// CFC twin of T_SafeConnShutdown_Tests: the same tests drawn as CFC diagrams, the way a TwinSAFE project is authored.
    FUNCTION_BLOCK T_SafeConnShutdown_Tests_CFC EXTENDS T_SafeCfcTestSuite
    VAR
    // Test_DeactivateShutsDownConnection
    group_1 : T_SafeGroup;
    conn_1 : T_SafeConnection(group := group_1);
    fb_1 : T_SafeConnShutdown(group := group_1, connection := conn_1);
END_VAR

Test_DeactivateShutsDownConnection();

METHOD PRIVATE Test_DeactivateShutsDownConnection
// note: this text did not pass the execution check against the stored diagram
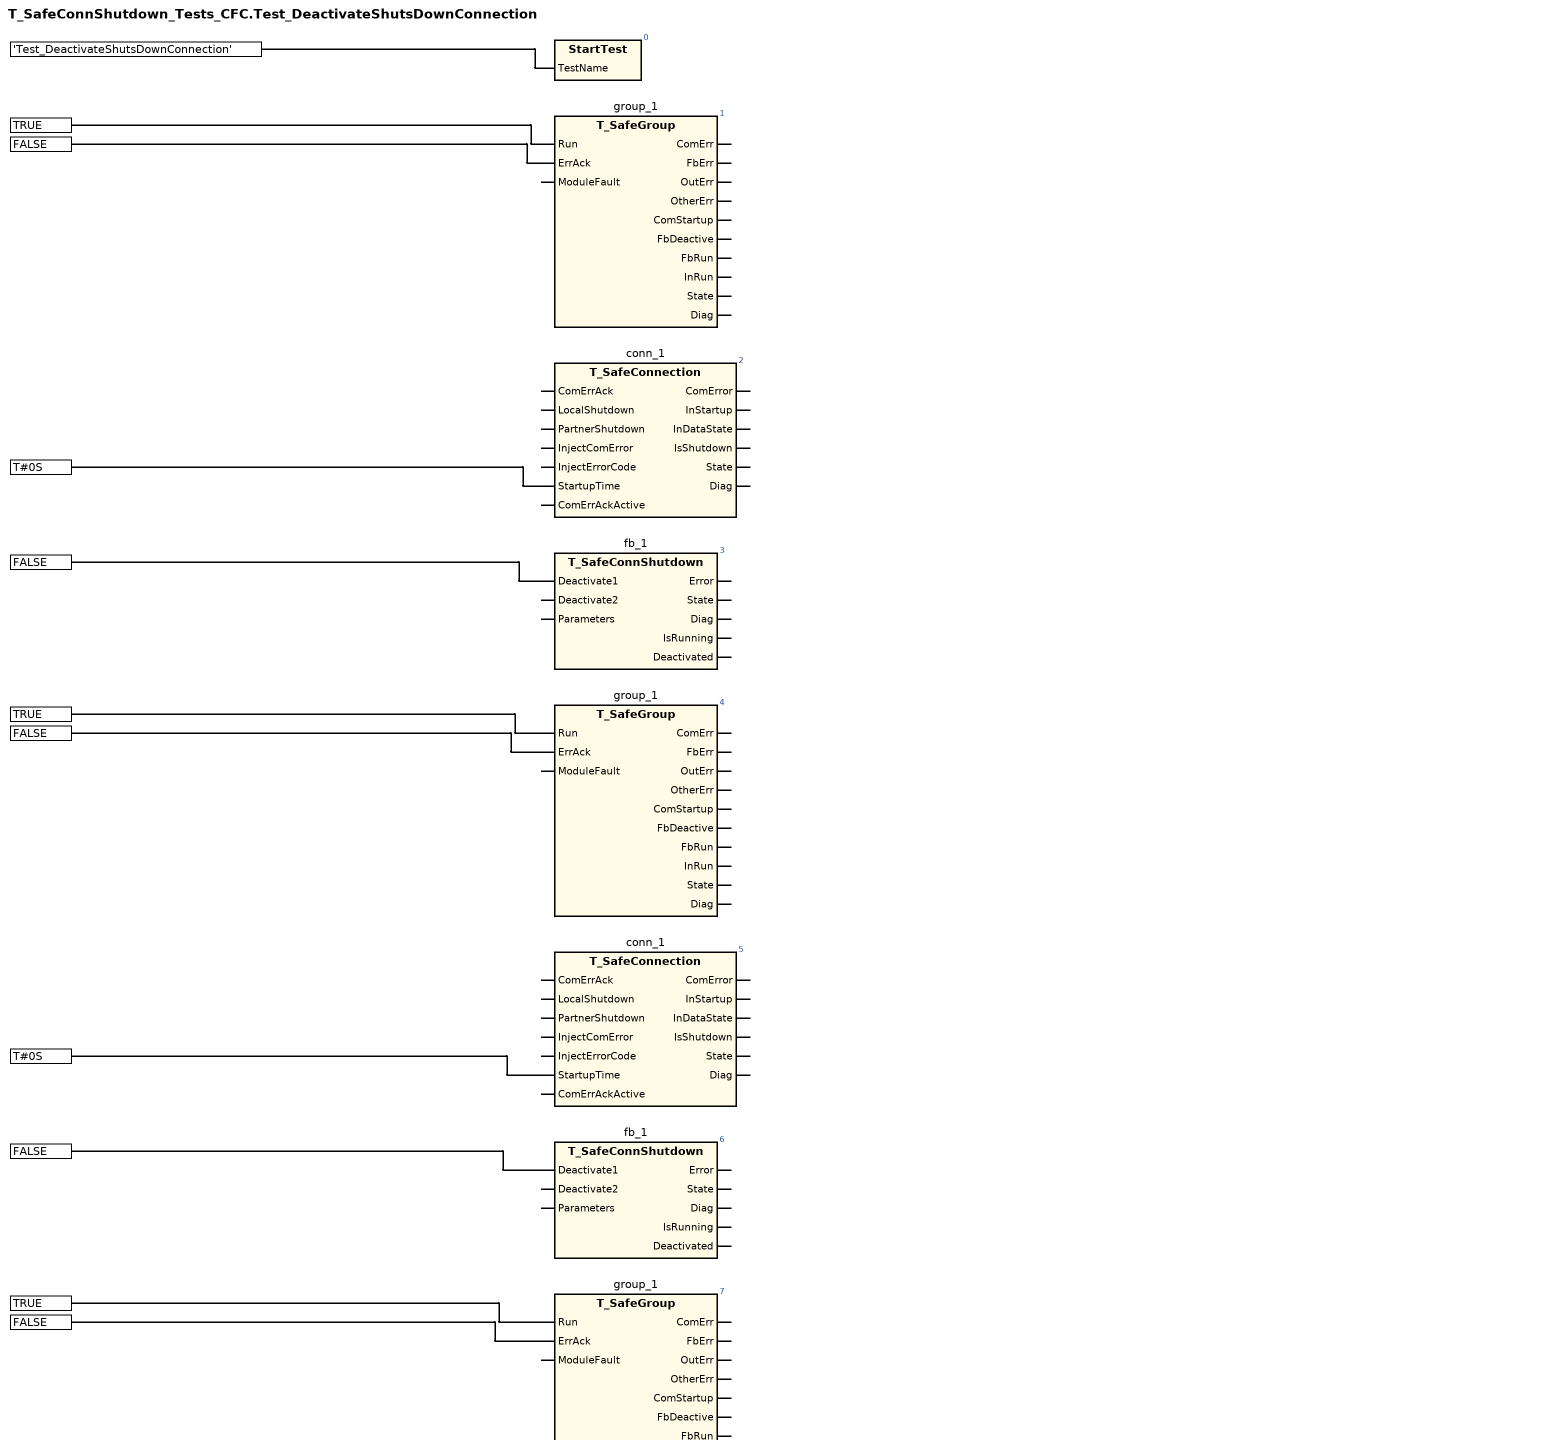
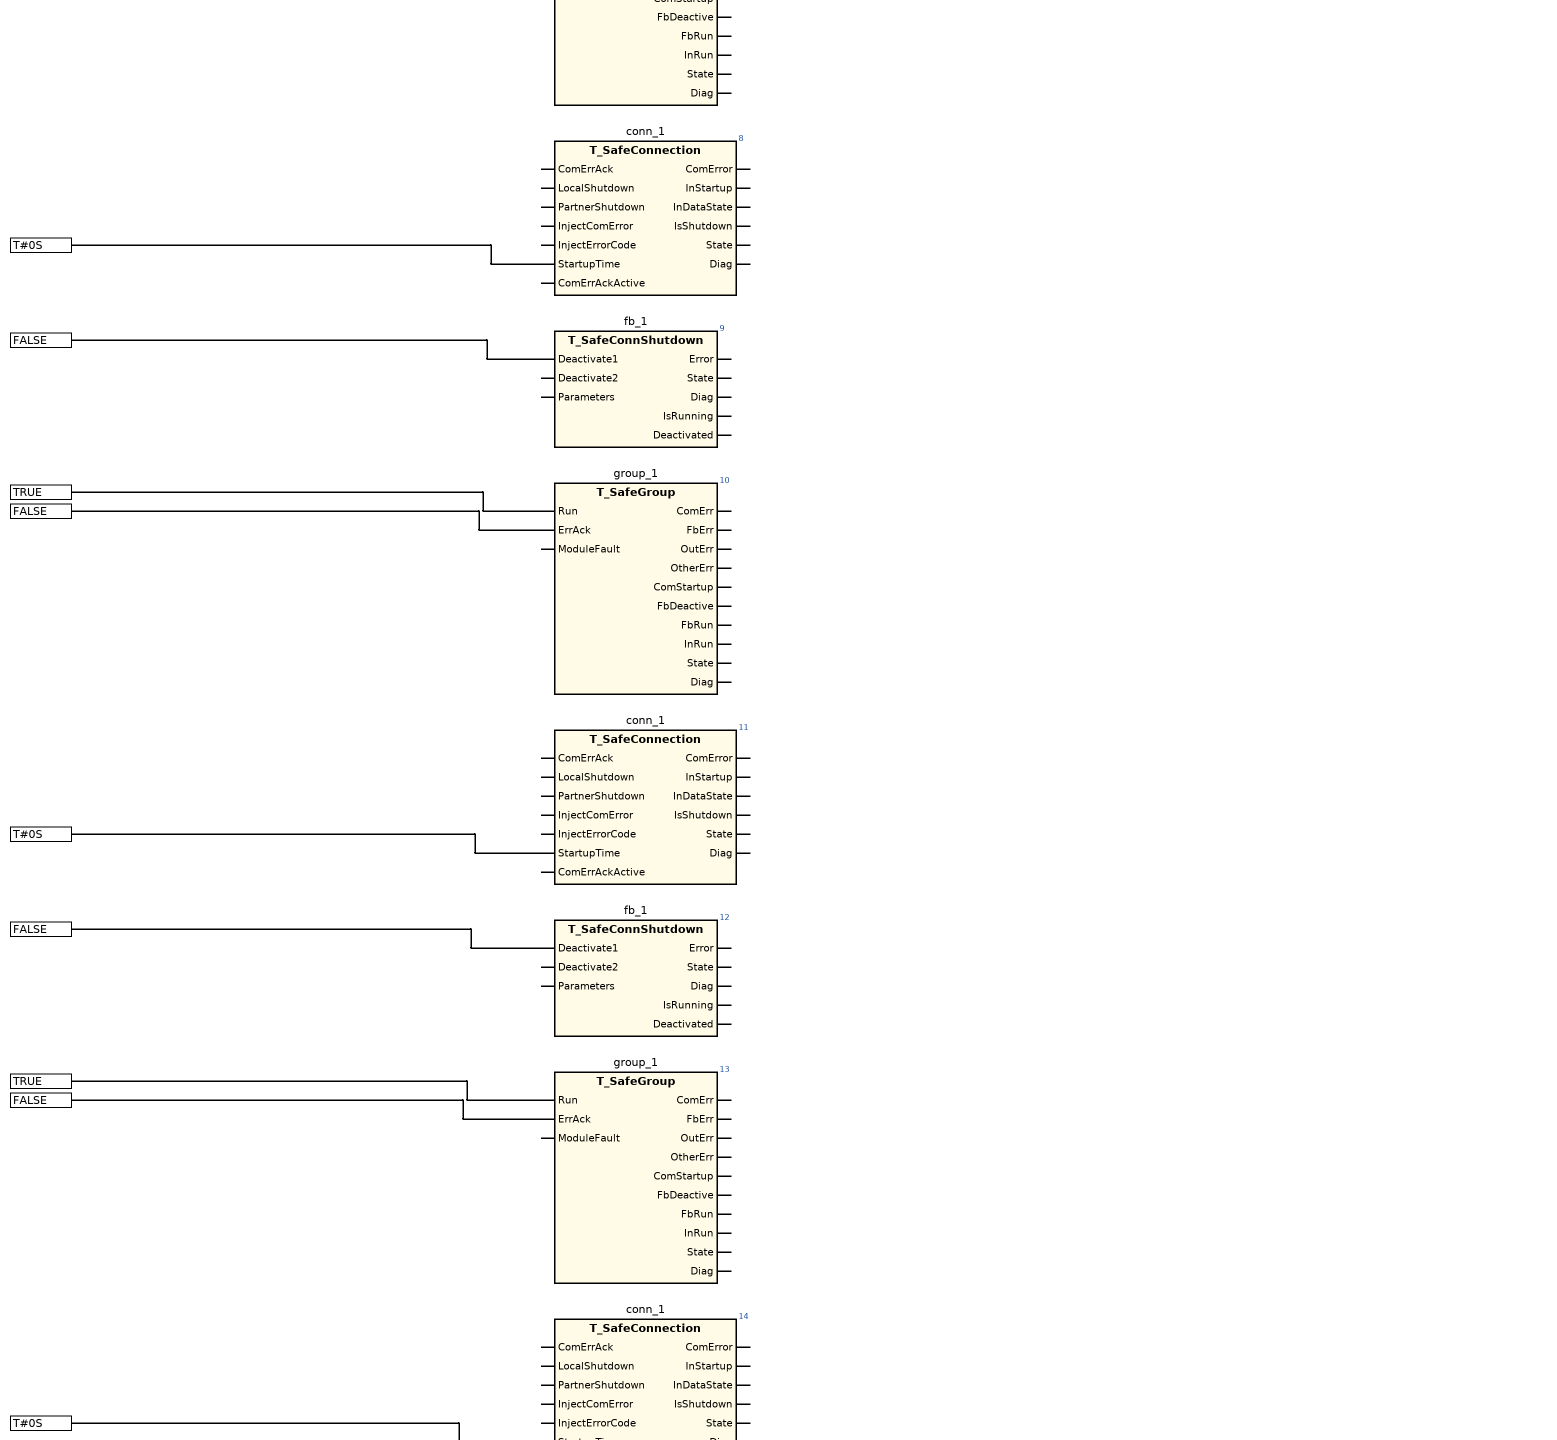
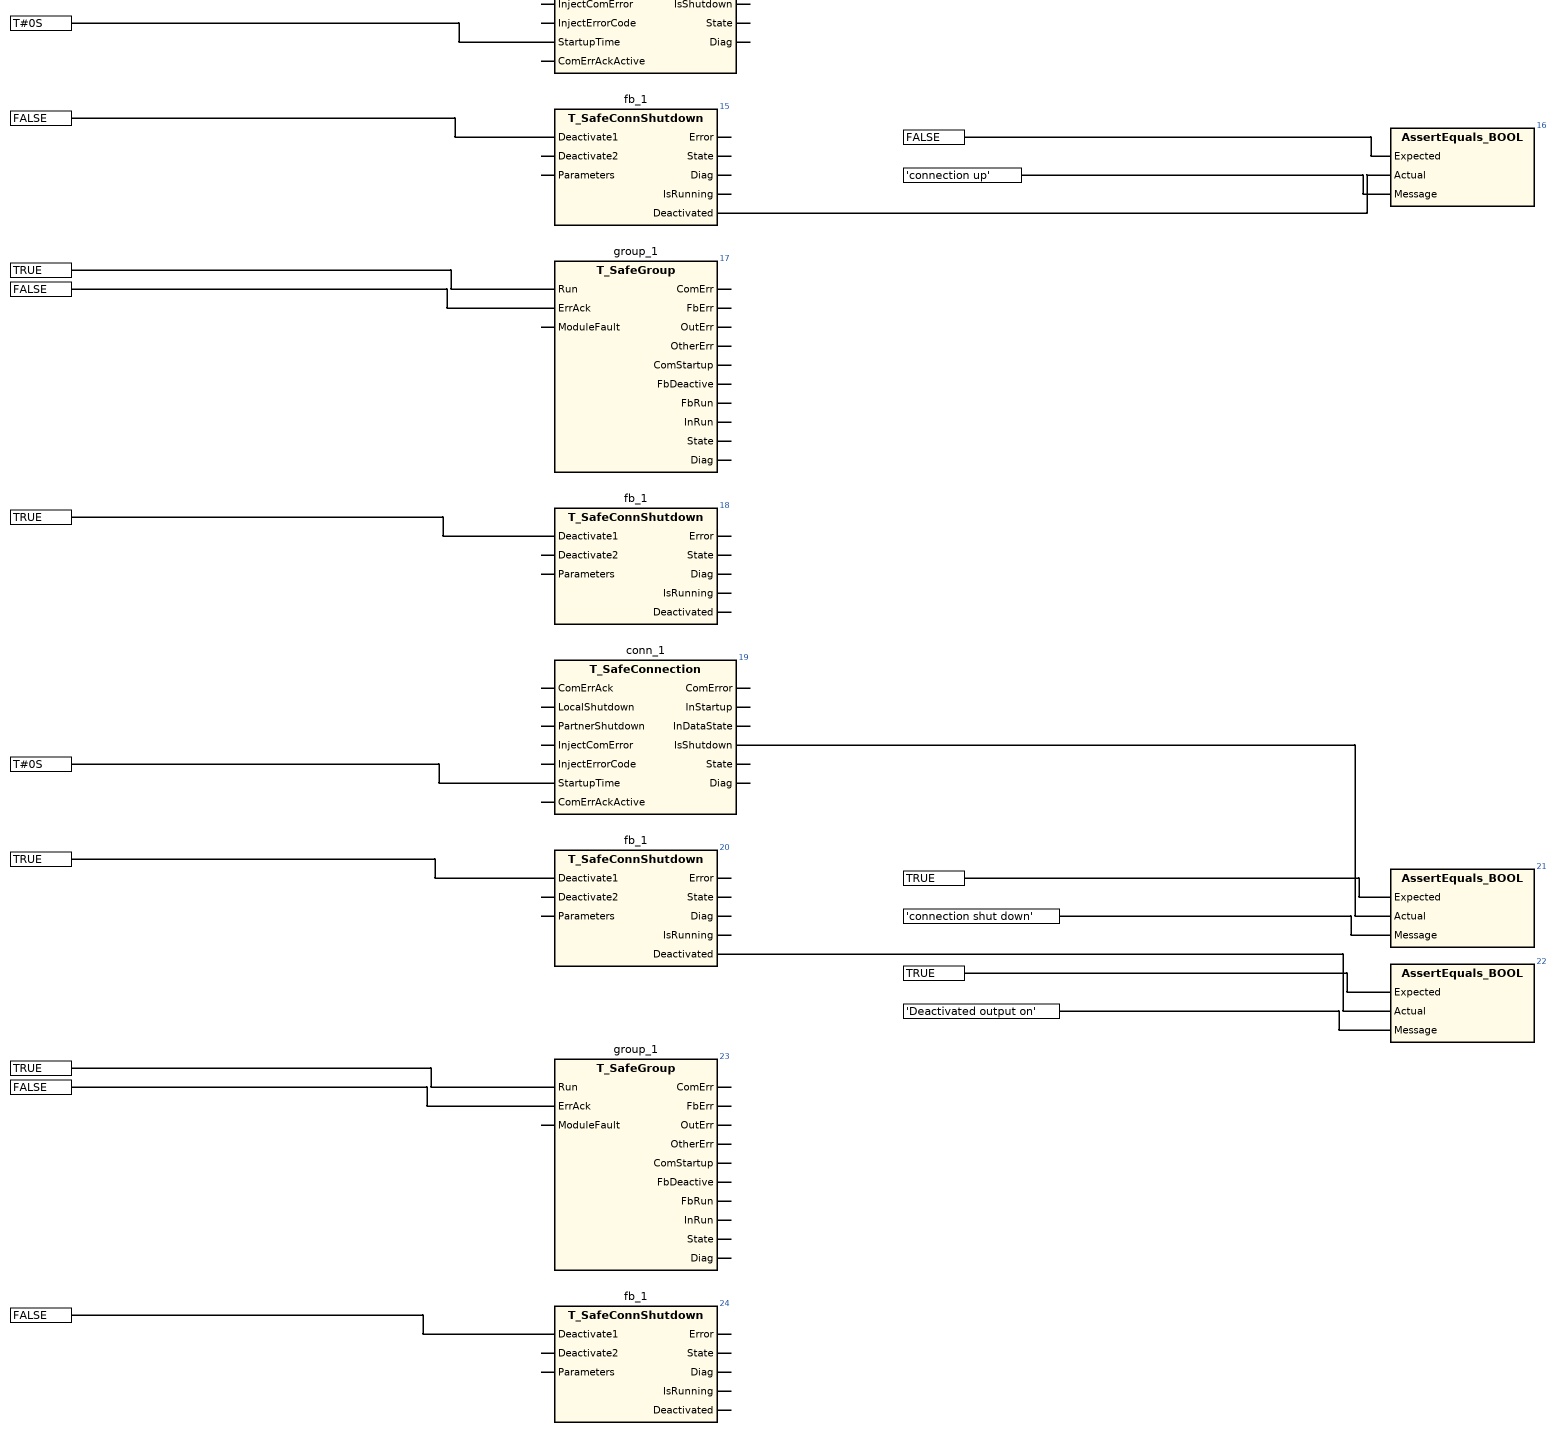
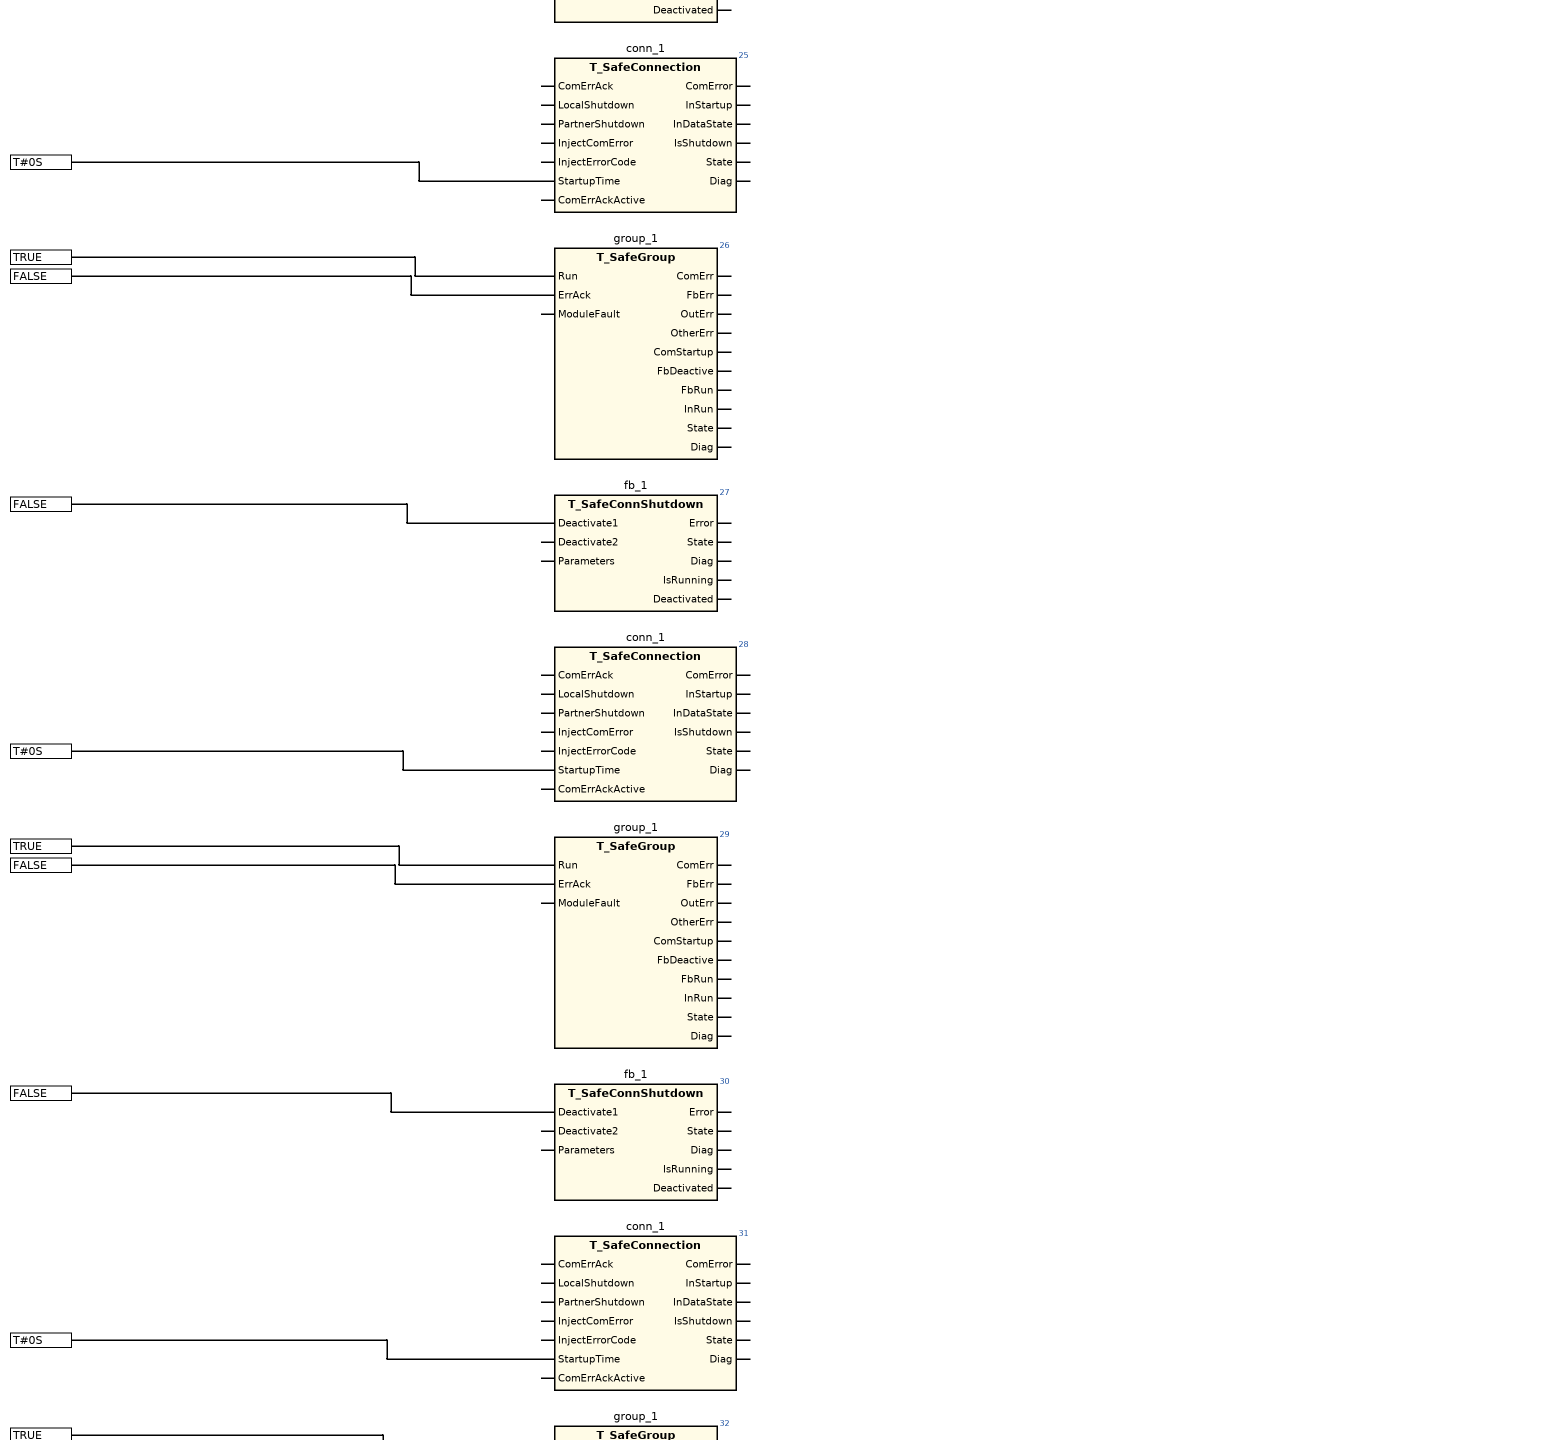
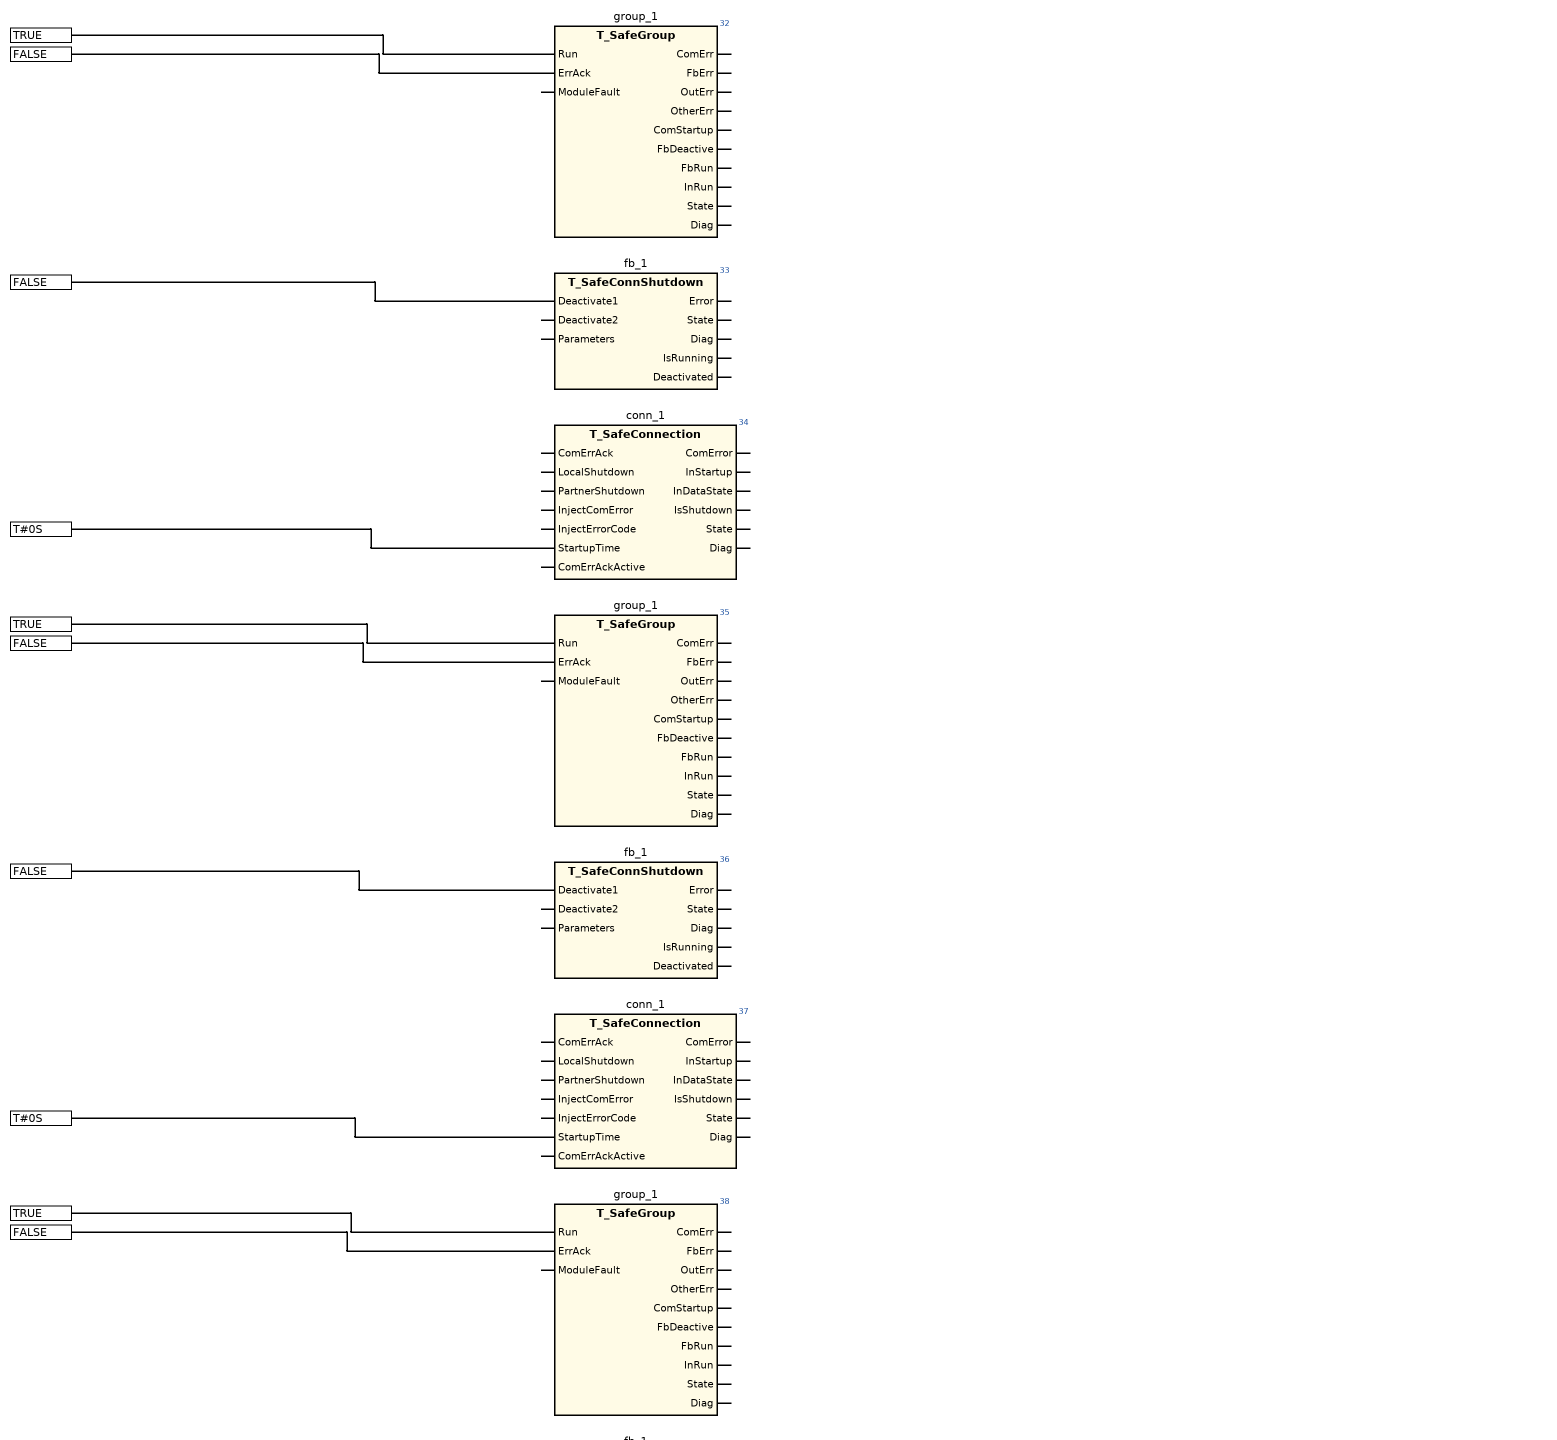
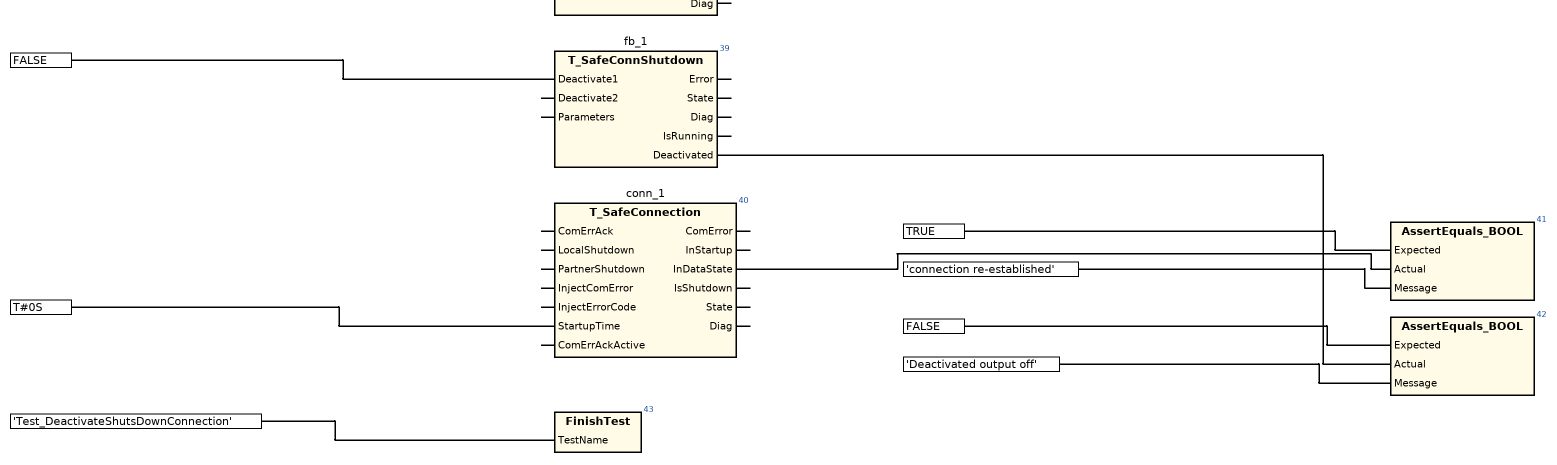
StartTest(TestName := 'Test_DeactivateShutsDownConnection');
group_1(Run := TRUE, ErrAck := FALSE); // T_SafeGroup
conn_1(StartupTime := T#0S); // T_SafeConnection
fb_1(Deactivate1 := FALSE); // T_SafeConnShutdown
group_1(Run := TRUE, ErrAck := FALSE); // T_SafeGroup
conn_1(StartupTime := T#0S); // T_SafeConnection
fb_1(Deactivate1 := FALSE); // T_SafeConnShutdown
group_1(Run := TRUE, ErrAck := FALSE); // T_SafeGroup
conn_1(StartupTime := T#0S); // T_SafeConnection
fb_1(Deactivate1 := FALSE); // T_SafeConnShutdown
group_1(Run := TRUE, ErrAck := FALSE); // T_SafeGroup
conn_1(StartupTime := T#0S); // T_SafeConnection
fb_1(Deactivate1 := FALSE); // T_SafeConnShutdown
group_1(Run := TRUE, ErrAck := FALSE); // T_SafeGroup
conn_1(StartupTime := T#0S); // T_SafeConnection
fb_1(Deactivate1 := FALSE); // T_SafeConnShutdown
AssertEquals_BOOL(Expected := FALSE, Actual := fb_1.Deactivated, Message := 'connection up');
group_1(Run := TRUE, ErrAck := FALSE); // T_SafeGroup
fb_1(Deactivate1 := TRUE); // T_SafeConnShutdown
conn_1(StartupTime := T#0S); // T_SafeConnection
fb_1(Deactivate1 := TRUE); // T_SafeConnShutdown
AssertEquals_BOOL(Expected := TRUE, Actual := conn_1.IsShutdown, Message := 'connection shut down');
AssertEquals_BOOL(Expected := TRUE, Actual := fb_1.Deactivated, Message := 'Deactivated output on');
group_1(Run := TRUE, ErrAck := FALSE); // T_SafeGroup
fb_1(Deactivate1 := FALSE); // T_SafeConnShutdown
conn_1(StartupTime := T#0S); // T_SafeConnection
group_1(Run := TRUE, ErrAck := FALSE); // T_SafeGroup
fb_1(Deactivate1 := FALSE); // T_SafeConnShutdown
conn_1(StartupTime := T#0S); // T_SafeConnection
group_1(Run := TRUE, ErrAck := FALSE); // T_SafeGroup
fb_1(Deactivate1 := FALSE); // T_SafeConnShutdown
conn_1(StartupTime := T#0S); // T_SafeConnection
group_1(Run := TRUE, ErrAck := FALSE); // T_SafeGroup
fb_1(Deactivate1 := FALSE); // T_SafeConnShutdown
conn_1(StartupTime := T#0S); // T_SafeConnection
group_1(Run := TRUE, ErrAck := FALSE); // T_SafeGroup
fb_1(Deactivate1 := FALSE); // T_SafeConnShutdown
conn_1(StartupTime := T#0S); // T_SafeConnection
group_1(Run := TRUE, ErrAck := FALSE); // T_SafeGroup
fb_1(Deactivate1 := FALSE); // T_SafeConnShutdown
conn_1(StartupTime := T#0S); // T_SafeConnection
AssertEquals_BOOL(Expected := TRUE, Actual := conn_1.InDataState, Message := 'connection re-established');
AssertEquals_BOOL(Expected := FALSE, Actual := fb_1.Deactivated, Message := 'Deactivated output off');
FinishTest(TestName := 'Test_DeactivateShutsDownConnection');
END_METHOD

END_FUNCTION_BLOCK

(* stored: Version 1.1.0.1, ProductVersion 3.1.4026.22
   POU T_SafeConnShutdown_Tests_CFC: Id {990feee4-9372-59d2-b479-6cfe606a9a7c}, SpecialFunc None
   Method Test_DeactivateShutsDownConnection: Id {44375d60-e47b-505d-9f4a-44c6bafc46e3} *)
